       5://SYSTEM 5
           "CNV_ID_HMI" := "Settings_DB".ECnv_Sys[5].ID; // EXTRACTOR CONVEYOR
           "CNV_HMI".CNV2_Selected[5] := "CNV2_Selected";
           CASE "CNV_Level_Selected" OF
               1: //LEVEL 1
                   IF "CNV2_Selected" = 1 THEN
                       "CNV_ID_HMI(1)" := "Settings_DB".LCnv_Sys[5].Cnv_Level[1].Cnv1.ID; //CNV 1
                   ELSIF "CNV2_Selected" = 2 THEN
                       "CNV_ID_HMI(1)" := "Settings_DB".LCnv_Sys[5].Cnv_Level[1].Cnv2.ID; //CNV 2
                   END_IF;
               2: //LEVEL 2
                   IF "CNV2_Selected" = 1 THEN
                       "CNV_ID_HMI(1)" := "Settings_DB".LCnv_Sys[5].Cnv_Level[2].Cnv1.ID; //CNV 1
                   ELSIF "CNV2_Selected" = 2 THEN
                       "CNV_ID_HMI(1)" := "Settings_DB".LCnv_Sys[5].Cnv_Level[2].Cnv2.ID; //CNV 2
                   END_IF;
               3: //LEVEL 3
                   IF "CNV2_Selected" = 1 THEN
                       "CNV_ID_HMI(1)" := "Settings_DB".LCnv_Sys[5].Cnv_Level[3].Cnv1.ID; //CNV 1
                   ELSIF "CNV2_Selected" = 2 THEN
                       "CNV_ID_HMI(1)" := "Settings_DB".LCnv_Sys[5].Cnv_Level[3].Cnv2.ID; //CNV 2
                   END_IF;
               4: //LEVEL 4
                   IF "CNV2_Selected" = 1 THEN
                       "CNV_ID_HMI(1)" := "Settings_DB".LCnv_Sys[5].Cnv_Level[4].Cnv1.ID; //CNV 1
                   ELSIF "CNV2_Selected" = 2 THEN
                       "CNV_ID_HMI(1)" := "Settings_DB".LCnv_Sys[5].Cnv_Level[4].Cnv2.ID; //CNV 2
                   END_IF;
               5: //LEVEL 5
                   IF "CNV2_Selected" = 1 THEN
                       "CNV_ID_HMI(1)" := "Settings_DB".LCnv_Sys[5].Cnv_Level[5].Cnv1.ID; //CNV 1
                   ELSIF "CNV2_Selected" = 2 THEN
                       "CNV_ID_HMI(1)" := "Settings_DB".LCnv_Sys[5].Cnv_Level[5].Cnv2.ID; //CNV 2
                   END_IF;
               6: //LEVEL 6
                   IF "CNV2_Selected" = 1 THEN
                       "CNV_ID_HMI(1)" := "Settings_DB".LCnv_Sys[5].Cnv_Level[6].Cnv1.ID; //CNV 1
                   ELSIF "CNV2_Selected" = 2 THEN
                       "CNV_ID_HMI(1)" := "Settings_DB".LCnv_Sys[5].Cnv_Level[6].Cnv2.ID; //CNV 2
                   END_IF;
               7: //LEVEL 7
                   IF "CNV2_Selected" = 1 THEN
                       "CNV_ID_HMI(1)" := "Settings_DB".LCnv_Sys[5].Cnv_Level[7].Cnv1.ID; //CNV 1
                   ELSIF "CNV2_Selected" = 2 THEN
                       "CNV_ID_HMI(1)" := "Settings_DB".LCnv_Sys[5].Cnv_Level[7].Cnv2.ID; //CNV 2
                   END_IF;
               8: //LEVEL 8
                   IF "CNV2_Selected" = 1 THEN
                       "CNV_ID_HMI(1)" := "Settings_DB".LCnv_Sys[5].Cnv_Level[8].Cnv1.ID; //CNV 1
                   ELSIF "CNV2_Selected" = 2 THEN
                       "CNV_ID_HMI(1)" := "Settings_DB".LCnv_Sys[5].Cnv_Level[8].Cnv2.ID; //CNV 2
                   END_IF;
           END_CASE;
   END_CASE;
END_FUNCTION

FUNCTION "CNV_Selector_1" : Void   // FC60, SCL
{ S7_Optimized_Access := 'TRUE' }
VERSION : 0.1
// stored: AutoNumber true, IsIECCheckEnabled false, SetENOAutomatically false, UDAEnableTagReadback false
   VAR_INPUT
      Sys_No : UInt;
      Zone : UInt;
      CNV1_2_Selected : UInt;
   END_VAR
   VAR_OUTPUT
      ID : DInt;
      "ID(1)" : DInt;
   END_VAR
BEGIN
   //CNV SCREEN SELECTION
   CASE #Sys_No OF
       0:
           #ID := 0;
           #"ID(1)" := 0;

       1://SYSTEM 1
           #ID := "Settings_DB".ECnv_Sys[1].ID; // EXTRACTOR CONVEYOR
           CASE #Zone OF
               11: //LEVEL 1
                   IF #CNV1_2_Selected = 1 THEN
                       #"ID(1)" := "Settings_DB".LCnv_Sys[1].Cnv_Level[1].Cnv1.ID; //CNV 1
                   ELSIF #CNV1_2_Selected = 2 THEN
                       #"ID(1)" := "Settings_DB".LCnv_Sys[1].Cnv_Level[1].Cnv2.ID; //CNV 2
                   END_IF;
               12: //LEVEL 2
                   IF #CNV1_2_Selected = 1 THEN
                       #"ID(1)" := "Settings_DB".LCnv_Sys[1].Cnv_Level[2].Cnv1.ID; //CNV 1
                   ELSIF #CNV1_2_Selected = 2 THEN
                       #"ID(1)" := "Settings_DB".LCnv_Sys[1].Cnv_Level[2].Cnv2.ID; //CNV 2
                   END_IF;
               13: //LEVEL 3
                   IF #CNV1_2_Selected = 1 THEN
                       #"ID(1)" := "Settings_DB".LCnv_Sys[1].Cnv_Level[3].Cnv1.ID; //CNV 1
                   ELSIF #CNV1_2_Selected = 2 THEN
                       #"ID(1)" := "Settings_DB".LCnv_Sys[1].Cnv_Level[3].Cnv2.ID; //CNV 2
                   END_IF;
               14: //LEVEL 4
                   IF #CNV1_2_Selected = 1 THEN
                       #"ID(1)" := "Settings_DB".LCnv_Sys[1].Cnv_Level[4].Cnv1.ID; //CNV 1
                   ELSIF #CNV1_2_Selected = 2 THEN
                       #"ID(1)" := "Settings_DB".LCnv_Sys[1].Cnv_Level[4].Cnv2.ID; //CNV 2
                   END_IF;
               15: //LEVEL 5
                   IF #CNV1_2_Selected = 1 THEN
                       #"ID(1)" := "Settings_DB".LCnv_Sys[1].Cnv_Level[5].Cnv1.ID; //CNV 1
                   ELSIF #CNV1_2_Selected = 2 THEN
                       #"ID(1)" := "Settings_DB".LCnv_Sys[1].Cnv_Level[5].Cnv2.ID; //CNV 2
                   END_IF;
               16: //LEVEL 6
                   IF #CNV1_2_Selected = 1 THEN
                       #"ID(1)" := "Settings_DB".LCnv_Sys[1].Cnv_Level[6].Cnv1.ID; //CNV 1
                   ELSIF #CNV1_2_Selected = 2 THEN
                       #"ID(1)" := "Settings_DB".LCnv_Sys[1].Cnv_Level[6].Cnv2.ID; //CNV 2
                   END_IF;
               17: //LEVEL 7
                   IF #CNV1_2_Selected = 1 THEN
                       #"ID(1)" := "Settings_DB".LCnv_Sys[1].Cnv_Level[7].Cnv1.ID; //CNV 1
                   ELSIF #CNV1_2_Selected = 2 THEN
                       #"ID(1)" := "Settings_DB".LCnv_Sys[1].Cnv_Level[7].Cnv2.ID; //CNV 2
                   END_IF;
               18: //LEVEL 8
                   IF #CNV1_2_Selected = 1 THEN
                       #"ID(1)" := "Settings_DB".LCnv_Sys[1].Cnv_Level[8].Cnv1.ID; //CNV 1
                   ELSIF #CNV1_2_Selected = 2 THEN
                       #"ID(1)" := "Settings_DB".LCnv_Sys[1].Cnv_Level[8].Cnv2.ID; //CNV 2
                   END_IF;
               19: //LEVEL 1
                   IF #CNV1_2_Selected = 1 THEN
                       #"ID(1)" := "Settings_DB".LCnv_Sys[1].Cnv_Level[1].Cnv1.ID; //CNV 1
                   ELSIF #CNV1_2_Selected = 2 THEN
                       #"ID(1)" := "Settings_DB".LCnv_Sys[1].Cnv_Level[1].Cnv2.ID; //CNV 2
                   END_IF;
           END_CASE;

       2://SYSTEM 2
           #ID := "Settings_DB".ECnv_Sys[2].ID; // EXTRACTOR CONVEYOR
           CASE #Zone OF
               21: //LEVEL 1
                   IF #CNV1_2_Selected = 1 THEN
                       #"ID(1)" := "Settings_DB".LCnv_Sys[2].Cnv_Level[1].Cnv1.ID; //CNV 1
                   ELSIF #CNV1_2_Selected = 2 THEN
                       #"ID(1)" := "Settings_DB".LCnv_Sys[2].Cnv_Level[1].Cnv2.ID; //CNV 2
                   END_IF;
               22: //LEVEL 2
                   IF #CNV1_2_Selected = 1 THEN
                       #"ID(1)" := "Settings_DB".LCnv_Sys[2].Cnv_Level[2].Cnv1.ID; //CNV 1
                   ELSIF #CNV1_2_Selected = 2 THEN
                       #"ID(1)" := "Settings_DB".LCnv_Sys[2].Cnv_Level[2].Cnv2.ID; //CNV 2
                   END_IF;
               23: //LEVEL 3
                   IF #CNV1_2_Selected = 1 THEN
                       #"ID(1)" := "Settings_DB".LCnv_Sys[2].Cnv_Level[3].Cnv1.ID; //CNV 1
                   ELSIF #CNV1_2_Selected = 2 THEN
                       #"ID(1)" := "Settings_DB".LCnv_Sys[2].Cnv_Level[3].Cnv2.ID; //CNV 2
                   END_IF;
               24: //LEVEL 4
                   IF #CNV1_2_Selected = 1 THEN
                       #"ID(1)" := "Settings_DB".LCnv_Sys[2].Cnv_Level[4].Cnv1.ID; //CNV 1
                   ELSIF #CNV1_2_Selected = 2 THEN
                       #"ID(1)" := "Settings_DB".LCnv_Sys[2].Cnv_Level[4].Cnv2.ID; //CNV 2
                   END_IF;
               25: //LEVEL 5
                   IF #CNV1_2_Selected = 1 THEN
                       #"ID(1)" := "Settings_DB".LCnv_Sys[2].Cnv_Level[5].Cnv1.ID; //CNV 1
                   ELSIF #CNV1_2_Selected = 2 THEN
                       #"ID(1)" := "Settings_DB".LCnv_Sys[2].Cnv_Level[5].Cnv2.ID; //CNV 2
                   END_IF;
               26: //LEVEL 6
                   IF #CNV1_2_Selected = 1 THEN
                       #"ID(1)" := "Settings_DB".LCnv_Sys[2].Cnv_Level[6].Cnv1.ID; //CNV 1
                   ELSIF #CNV1_2_Selected = 2 THEN
                       #"ID(1)" := "Settings_DB".LCnv_Sys[2].Cnv_Level[6].Cnv2.ID; //CNV 2
                   END_IF;
               27: //LEVEL 7
                   IF #CNV1_2_Selected = 1 THEN
                       #"ID(1)" := "Settings_DB".LCnv_Sys[2].Cnv_Level[7].Cnv1.ID; //CNV 1
                   ELSIF #CNV1_2_Selected = 2 THEN
                       #"ID(1)" := "Settings_DB".LCnv_Sys[2].Cnv_Level[7].Cnv2.ID; //CNV 2
                   END_IF;
               28: //LEVEL 8
                   IF #CNV1_2_Selected = 1 THEN
                       #"ID(1)" := "Settings_DB".LCnv_Sys[2].Cnv_Level[8].Cnv1.ID; //CNV 1
                   ELSIF #CNV1_2_Selected = 2 THEN
                       #"ID(1)" := "Settings_DB".LCnv_Sys[2].Cnv_Level[8].Cnv2.ID; //CNV 2
                   END_IF;
               29: //LEVEL 1
                   IF #CNV1_2_Selected = 1 THEN
                       #"ID(1)" := "Settings_DB".LCnv_Sys[2].Cnv_Level[1].Cnv1.ID; //CNV 1
                   ELSIF #CNV1_2_Selected = 2 THEN
                       #"ID(1)" := "Settings_DB".LCnv_Sys[2].Cnv_Level[1].Cnv2.ID; //CNV 2
                   END_IF;
           END_CASE;

       3://SYSTEM 3
           #ID := "Settings_DB".ECnv_Sys[3].ID; // EXTRACTOR CONVEYOR
           CASE #Zone OF
               31: //LEVEL 1
                   IF #CNV1_2_Selected = 1 THEN
                       #"ID(1)" := "Settings_DB".LCnv_Sys[3].Cnv_Level[1].Cnv1.ID; //CNV 1
                   ELSIF #CNV1_2_Selected = 2 THEN
                       #"ID(1)" := "Settings_DB".LCnv_Sys[3].Cnv_Level[1].Cnv2.ID; //CNV 2
                   END_IF;
               32: //LEVEL 2
                   IF #CNV1_2_Selected = 1 THEN
                       #"ID(1)" := "Settings_DB".LCnv_Sys[3].Cnv_Level[2].Cnv1.ID; //CNV 1
                   ELSIF #CNV1_2_Selected = 2 THEN
                       #"ID(1)" := "Settings_DB".LCnv_Sys[3].Cnv_Level[2].Cnv2.ID; //CNV 2
                   END_IF;
               33: //LEVEL 3
                   IF #CNV1_2_Selected = 1 THEN
                       #"ID(1)" := "Settings_DB".LCnv_Sys[3].Cnv_Level[3].Cnv1.ID; //CNV 1
                   ELSIF #CNV1_2_Selected = 2 THEN
                       #"ID(1)" := "Settings_DB".LCnv_Sys[3].Cnv_Level[3].Cnv2.ID; //CNV 2
                   END_IF;
               34: //LEVEL 4
                   IF #CNV1_2_Selected = 1 THEN
                       #"ID(1)" := "Settings_DB".LCnv_Sys[3].Cnv_Level[4].Cnv1.ID; //CNV 1
                   ELSIF #CNV1_2_Selected = 2 THEN
                       #"ID(1)" := "Settings_DB".LCnv_Sys[3].Cnv_Level[4].Cnv2.ID; //CNV 2
                   END_IF;
               35: //LEVEL 5
                   IF #CNV1_2_Selected = 1 THEN
                       #"ID(1)" := "Settings_DB".LCnv_Sys[3].Cnv_Level[5].Cnv1.ID; //CNV 1
                   ELSIF #CNV1_2_Selected = 2 THEN
                       #"ID(1)" := "Settings_DB".LCnv_Sys[3].Cnv_Level[5].Cnv2.ID; //CNV 2
                   END_IF;
               36: //LEVEL 6
                   IF #CNV1_2_Selected = 1 THEN
                       #"ID(1)" := "Settings_DB".LCnv_Sys[3].Cnv_Level[6].Cnv1.ID; //CNV 1
                   ELSIF #CNV1_2_Selected = 2 THEN
                       #"ID(1)" := "Settings_DB".LCnv_Sys[3].Cnv_Level[6].Cnv2.ID; //CNV 2
                   END_IF;
               37: //LEVEL 7
                   IF #CNV1_2_Selected = 1 THEN
                       #"ID(1)" := "Settings_DB".LCnv_Sys[3].Cnv_Level[7].Cnv1.ID; //CNV 1
                   ELSIF #CNV1_2_Selected = 2 THEN
                       #"ID(1)" := "Settings_DB".LCnv_Sys[3].Cnv_Level[7].Cnv2.ID; //CNV 2
                   END_IF;
               38: //LEVEL 8
                   IF #CNV1_2_Selected = 1 THEN
                       #"ID(1)" := "Settings_DB".LCnv_Sys[3].Cnv_Level[8].Cnv1.ID; //CNV 1
                   ELSIF #CNV1_2_Selected = 2 THEN
                       #"ID(1)" := "Settings_DB".LCnv_Sys[3].Cnv_Level[8].Cnv2.ID; //CNV 2
                   END_IF;
               39: //LEVEL 1
                   IF #CNV1_2_Selected = 1 THEN
                       #"ID(1)" := "Settings_DB".LCnv_Sys[3].Cnv_Level[1].Cnv1.ID; //CNV 1
                   ELSIF #CNV1_2_Selected = 2 THEN
                       #"ID(1)" := "Settings_DB".LCnv_Sys[3].Cnv_Level[1].Cnv2.ID; //CNV 2
                   END_IF;
           END_CASE;

       4://SYSTEM 4
           #ID := "Settings_DB".ECnv_Sys[4].ID; // EXTRACTOR CONVEYOR
           CASE #Zone OF
               41: //LEVEL 1
                   IF #CNV1_2_Selected = 1 THEN
                       #"ID(1)" := "Settings_DB".LCnv_Sys[4].Cnv_Level[1].Cnv1.ID; //CNV 1
                   ELSIF #CNV1_2_Selected = 2 THEN
                       #"ID(1)" := "Settings_DB".LCnv_Sys[4].Cnv_Level[1].Cnv2.ID; //CNV 2
                   END_IF;
               42: //LEVEL 2
                   IF #CNV1_2_Selected = 1 THEN
                       #"ID(1)" := "Settings_DB".LCnv_Sys[4].Cnv_Level[2].Cnv1.ID; //CNV 1
                   ELSIF #CNV1_2_Selected = 2 THEN
                       #"ID(1)" := "Settings_DB".LCnv_Sys[4].Cnv_Level[2].Cnv2.ID; //CNV 2
                   END_IF;
               43: //LEVEL 3
                   IF #CNV1_2_Selected = 1 THEN
                       #"ID(1)" := "Settings_DB".LCnv_Sys[4].Cnv_Level[3].Cnv1.ID; //CNV 1
                   ELSIF #CNV1_2_Selected = 2 THEN
                       #"ID(1)" := "Settings_DB".LCnv_Sys[4].Cnv_Level[3].Cnv2.ID; //CNV 2
                   END_IF;
               44: //LEVEL 4
                   IF #CNV1_2_Selected = 1 THEN
                       #"ID(1)" := "Settings_DB".LCnv_Sys[4].Cnv_Level[4].Cnv1.ID; //CNV 1
                   ELSIF #CNV1_2_Selected = 2 THEN
                       #"ID(1)" := "Settings_DB".LCnv_Sys[4].Cnv_Level[4].Cnv2.ID; //CNV 2
                   END_IF;
               45: //LEVEL 5
                   IF #CNV1_2_Selected = 1 THEN
                       #"ID(1)" := "Settings_DB".LCnv_Sys[4].Cnv_Level[5].Cnv1.ID; //CNV 1
                   ELSIF #CNV1_2_Selected = 2 THEN
                       #"ID(1)" := "Settings_DB".LCnv_Sys[4].Cnv_Level[5].Cnv2.ID; //CNV 2
                   END_IF;
               46: //LEVEL 6
                   IF #CNV1_2_Selected = 1 THEN
                       #"ID(1)" := "Settings_DB".LCnv_Sys[4].Cnv_Level[6].Cnv1.ID; //CNV 1
                   ELSIF #CNV1_2_Selected = 2 THEN
                       #"ID(1)" := "Settings_DB".LCnv_Sys[4].Cnv_Level[6].Cnv2.ID; //CNV 2
                   END_IF;
               47: //LEVEL 7
                   IF #CNV1_2_Selected = 1 THEN
                       #"ID(1)" := "Settings_DB".LCnv_Sys[4].Cnv_Level[7].Cnv1.ID; //CNV 1
                   ELSIF #CNV1_2_Selected = 2 THEN
                       #"ID(1)" := "Settings_DB".LCnv_Sys[4].Cnv_Level[7].Cnv2.ID; //CNV 2
                   END_IF;
               48: //LEVEL 8
                   IF #CNV1_2_Selected = 1 THEN
                       #"ID(1)" := "Settings_DB".LCnv_Sys[4].Cnv_Level[8].Cnv1.ID; //CNV 1
                   ELSIF #CNV1_2_Selected = 2 THEN
                       #"ID(1)" := "Settings_DB".LCnv_Sys[4].Cnv_Level[8].Cnv2.ID; //CNV 2
                   END_IF;
               49: //LEVEL 1
                   IF #CNV1_2_Selected = 1 THEN
                       #"ID(1)" := "Settings_DB".LCnv_Sys[4].Cnv_Level[1].Cnv1.ID; //CNV 1
                   ELSIF #CNV1_2_Selected = 2 THEN
                       #"ID(1)" := "Settings_DB".LCnv_Sys[4].Cnv_Level[1].Cnv2.ID; //CNV 2
                   END_IF;
           END_CASE;

       5://SYSTEM 5
           #ID := "Settings_DB".ECnv_Sys[5].ID; // EXTRACTOR CONVEYOR
           CASE #Zone OF
               51: //LEVEL 1
                   IF #CNV1_2_Selected = 1 THEN
                       #"ID(1)" := "Settings_DB".LCnv_Sys[5].Cnv_Level[1].Cnv1.ID; //CNV 1
                   ELSIF #CNV1_2_Selected = 2 THEN
                       #"ID(1)" := "Settings_DB".LCnv_Sys[5].Cnv_Level[1].Cnv2.ID; //CNV 2
                   END_IF;
               52: //LEVEL 2
                   IF #CNV1_2_Selected = 1 THEN
                       #"ID(1)" := "Settings_DB".LCnv_Sys[5].Cnv_Level[2].Cnv1.ID; //CNV 1
                   ELSIF #CNV1_2_Selected = 2 THEN
                       #"ID(1)" := "Settings_DB".LCnv_Sys[5].Cnv_Level[2].Cnv2.ID; //CNV 2
                   END_IF;
               53: //LEVEL 3
                   IF #CNV1_2_Selected = 1 THEN
                       #"ID(1)" := "Settings_DB".LCnv_Sys[5].Cnv_Level[3].Cnv1.ID; //CNV 1
                   ELSIF #CNV1_2_Selected = 2 THEN
                       #"ID(1)" := "Settings_DB".LCnv_Sys[5].Cnv_Level[3].Cnv2.ID; //CNV 2
                   END_IF;
               54: //LEVEL 4
                   IF #CNV1_2_Selected = 1 THEN
                       #"ID(1)" := "Settings_DB".LCnv_Sys[5].Cnv_Level[4].Cnv1.ID; //CNV 1
                   ELSIF #CNV1_2_Selected = 2 THEN
                       #"ID(1)" := "Settings_DB".LCnv_Sys[5].Cnv_Level[4].Cnv2.ID; //CNV 2
                   END_IF;
               55: //LEVEL 5
                   IF #CNV1_2_Selected = 1 THEN
                       #"ID(1)" := "Settings_DB".LCnv_Sys[5].Cnv_Level[5].Cnv1.ID; //CNV 1
                   ELSIF #CNV1_2_Selected = 2 THEN
                       #"ID(1)" := "Settings_DB".LCnv_Sys[5].Cnv_Level[5].Cnv2.ID; //CNV 2
                   END_IF;
               56: //LEVEL 6
                   IF #CNV1_2_Selected = 1 THEN
                       #"ID(1)" := "Settings_DB".LCnv_Sys[5].Cnv_Level[6].Cnv1.ID; //CNV 1
                   ELSIF #CNV1_2_Selected = 2 THEN
                       #"ID(1)" := "Settings_DB".LCnv_Sys[5].Cnv_Level[6].Cnv2.ID; //CNV 2
                   END_IF;
               57: //LEVEL 7
                   IF #CNV1_2_Selected = 1 THEN
                       #"ID(1)" := "Settings_DB".LCnv_Sys[5].Cnv_Level[7].Cnv1.ID; //CNV 1
                   ELSIF #CNV1_2_Selected = 2 THEN
                       #"ID(1)" := "Settings_DB".LCnv_Sys[5].Cnv_Level[7].Cnv2.ID; //CNV 2
                   END_IF;
               58: //LEVEL 8
                   IF #CNV1_2_Selected = 1 THEN
                       #"ID(1)" := "Settings_DB".LCnv_Sys[5].Cnv_Level[8].Cnv1.ID; //CNV 1
                   ELSIF #CNV1_2_Selected = 2 THEN
                       #"ID(1)" := "Settings_DB".LCnv_Sys[5].Cnv_Level[8].Cnv2.ID; //CNV 2
                   END_IF;
               59: //LEVEL 1
                   IF #CNV1_2_Selected = 1 THEN
                       #"ID(1)" := "Settings_DB".LCnv_Sys[5].Cnv_Level[1].Cnv1.ID; //CNV 1
                   ELSIF #CNV1_2_Selected = 2 THEN
                       #"ID(1)" := "Settings_DB".LCnv_Sys[5].Cnv_Level[1].Cnv2.ID; //CNV 2
                   END_IF;
           END_CASE;
   END_CASE;
END_FUNCTION

FUNCTION "CharsArrayToString" : String   // FC27, SCL
{ S7_Optimized_Access := 'TRUE' }
VERSION : 0.1
// stored: AutoNumber true, IsIECCheckEnabled false, SetENOAutomatically false, UDAEnableTagReadback false
   VAR_INPUT
      Lenght : Int;
      CharsArray : Array[1..16] of Char;
   END_VAR
   VAR_TEMP
      tempStr_1 : String;
      foundPos : Int;
      i : Int;
   END_VAR
BEGIN
   #tempStr_1 := '';
   FOR #i := 1 TO MIN(IN1 := #Lenght - 1, IN2 := 16) DO
       IF #CharsArray[#i] <> '$00' THEN
           #tempStr_1 := CONCAT(IN1 := #tempStr_1, IN2 := CHAR_TO_STRING(#CharsArray[#i]));
       END_IF;
   END_FOR;

   // Remove '$00'
   // string 1
   #foundPos := FIND(IN1 := #tempStr_1, IN2 := '$00');
   WHILE #foundPos > 0 DO
       #tempStr_1 := REPLACE(IN1 := #tempStr_1, IN2 := '', P := #foundPos, L := 1);
       #foundPos := FIND(IN1 := #tempStr_1, IN2 := '$00');
   END_WHILE;

   #CharsArrayToString := #tempStr_1;
END_FUNCTION

FUNCTION_BLOCK "Conveyor_HMI_FB"   // FB20, SCL
{ S7_Optimized_Access := 'TRUE' }
VERSION : 0.1
// stored: AutoNumber true, IsIECCheckEnabled false, IsRetainMemResEnabled false, MemoryReserve 100, SetENOAutomatically false, UDAEnableTagReadback false
   VAR
      R_Charge_Cnv_Commands { S7_SetPoint := 'True'} : R_TRIG;
      T_Reset_Charge { S7_SetPoint := 'True'} : TON_TIME;
   END_VAR
   VAR_TEMP
      i : UInt;
      J : UInt;
      No_Light_Guard : Bool;
   END_VAR
BEGIN
   "CNV_Selector"();

   REGION SEND/RECEIVE BUTTON
       IF "CNV_System_Selected" = 1 AND NOT "Control_DB".VTD_Sys[1].Running AND "Control_DB".VTD_Sys[1].Current_Level <> 0 THEN
           IF "CNV2_Selected" = 1 AND "HMI_DB".ScreenNo_Main = 2 THEN
               //CNV 1
               IF "Control_DB".ECnv_Sys[1].Cnv_Occupied AND NOT "Control_DB".LCnv_Sys[1].Cnv_Level["Control_DB".VTD_Sys[1].Current_Level].Cnv1.Cnv_Occupied AND
                   NOT "Control_DB".ECnv_Sys[1].Running AND NOT "Control_DB".LCnv_Sys[1].Cnv_Level["Control_DB".VTD_Sys[1].Current_Level].Cnv1.Running AND
                   "Control_DB".LCnv_Sys[1].Cnv_Level["Control_DB".VTD_Sys[1].Current_Level].Cnv1.Pallet_Type <> 1 AND "Control_DB".ECnv_Sys[1].Pallet_Type <> 5 THEN
                   "CNV_HMI".In_Out[1] := TRUE;
                   "CNV_In_Out" := TRUE;
               ELSIF NOT "Control_DB".ECnv_Sys[1].Cnv_Occupied AND "Control_DB".LCnv_Sys[1].Cnv_Level["Control_DB".VTD_Sys[1].Current_Level].Cnv1.Cnv_Occupied AND
                   NOT "Control_DB".ECnv_Sys[1].Running AND NOT "Control_DB".LCnv_Sys[1].Cnv_Level["Control_DB".VTD_Sys[1].Current_Level].Cnv1.Running THEN
                   "CNV_HMI".In_Out[1] := FALSE;
                   "CNV_In_Out" := FALSE;
               ELSE
                   ;
               END_IF;
               //CNV 2
           ELSIF "CNV2_Selected" = 2 AND "HMI_DB".ScreenNo_Main = 2 THEN   //CNV 2
               IF "Control_DB".ECnv_Sys[1].Cnv_Occupied AND NOT "Control_DB".LCnv_Sys[1].Cnv_Level["Control_DB".VTD_Sys[1].Current_Level].Cnv2.Cnv_Occupied AND
                   NOT "Control_DB".ECnv_Sys[1].Running AND NOT "Control_DB".LCnv_Sys[1].Cnv_Level["Control_DB".VTD_Sys[1].Current_Level].Cnv2.Running AND
                   "Control_DB".LCnv_Sys[1].Cnv_Level["Control_DB".VTD_Sys[1].Current_Level].Cnv2.Pallet_Type <> 1 AND "Control_DB".ECnv_Sys[1].Pallet_Type <> 5 THEN
                   "CNV_HMI".In_Out[1] := TRUE;
                   "CNV_In_Out" := TRUE;
               ELSIF NOT "Control_DB".ECnv_Sys[1].Cnv_Occupied AND "Control_DB".LCnv_Sys[1].Cnv_Level["Control_DB".VTD_Sys[1].Current_Level].Cnv2.Cnv_Occupied AND
                   NOT "Control_DB".ECnv_Sys[1].Running AND NOT "Control_DB".LCnv_Sys[1].Cnv_Level["Control_DB".VTD_Sys[1].Current_Level].Cnv2.Running THEN
                   "CNV_HMI".In_Out[1] := FALSE;
                   "CNV_In_Out" := FALSE;
               ELSE
                   ;
               END_IF;
           END_IF;
       END_IF;

       IF "CNV_System_Selected" = 2 AND NOT "Control_DB".VTD_Sys[2].Running AND "Control_DB".VTD_Sys[2].Current_Level <> 0 THEN
           IF "CNV2_Selected" = 1 AND "HMI_DB".ScreenNo_Main = 2 THEN
               //CNV 1
               IF "Control_DB".ECnv_Sys[2].Cnv_Occupied AND NOT "Control_DB".LCnv_Sys[2].Cnv_Level["Control_DB".VTD_Sys[2].Current_Level].Cnv1.Cnv_Occupied AND
                   NOT "Control_DB".ECnv_Sys[2].Running AND NOT "Control_DB".LCnv_Sys[2].Cnv_Level["Control_DB".VTD_Sys[2].Current_Level].Cnv1.Running AND
                   "Control_DB".LCnv_Sys[2].Cnv_Level["Control_DB".VTD_Sys[2].Current_Level].Cnv1.Pallet_Type <> 1 AND "Control_DB".ECnv_Sys[2].Pallet_Type <> 5 THEN
                   "CNV_HMI".In_Out[2] := TRUE;
                   "CNV_In_Out" := TRUE;
               ELSIF NOT "Control_DB".ECnv_Sys[2].Cnv_Occupied AND "Control_DB".LCnv_Sys[2].Cnv_Level["Control_DB".VTD_Sys[2].Current_Level].Cnv1.Cnv_Occupied AND
                   NOT "Control_DB".ECnv_Sys[2].Running AND NOT "Control_DB".LCnv_Sys[2].Cnv_Level["Control_DB".VTD_Sys[2].Current_Level].Cnv1.Running THEN
                   "CNV_HMI".In_Out[2] := FALSE;
                   "CNV_In_Out" := FALSE;
               ELSE
                   ;
               END_IF;
               //CNV 2
           ELSIF "CNV2_Selected" = 2 AND "HMI_DB".ScreenNo_Main = 2 THEN   //CNV 2
               IF "Control_DB".ECnv_Sys[2].Cnv_Occupied AND NOT "Control_DB".LCnv_Sys[2].Cnv_Level["Control_DB".VTD_Sys[2].Current_Level].Cnv2.Cnv_Occupied AND
                   NOT "Control_DB".ECnv_Sys[2].Running AND NOT "Control_DB".LCnv_Sys[2].Cnv_Level["Control_DB".VTD_Sys[2].Current_Level].Cnv2.Running AND
                   "Control_DB".LCnv_Sys[2].Cnv_Level["Control_DB".VTD_Sys[2].Current_Level].Cnv2.Pallet_Type <> 1 AND "Control_DB".ECnv_Sys[2].Pallet_Type <> 5 THEN
                   "CNV_HMI".In_Out[2] := TRUE;
                   "CNV_In_Out" := TRUE;
               ELSIF NOT "Control_DB".ECnv_Sys[2].Cnv_Occupied AND "Control_DB".LCnv_Sys[2].Cnv_Level["Control_DB".VTD_Sys[2].Current_Level].Cnv2.Cnv_Occupied AND
                   NOT "Control_DB".ECnv_Sys[2].Running AND NOT "Control_DB".LCnv_Sys[2].Cnv_Level["Control_DB".VTD_Sys[2].Current_Level].Cnv2.Running THEN
                   "CNV_HMI".In_Out[2] := FALSE;
                   "CNV_In_Out" := FALSE;
               ELSE
                   ;
               END_IF;
           END_IF;
       END_IF;

       IF "CNV_System_Selected" = 3 AND NOT "Control_DB".VTD_Sys[3].Running AND "Control_DB".VTD_Sys[3].Current_Level <> 0 THEN
           IF "CNV2_Selected" = 1 AND "HMI_DB".ScreenNo_Main = 2 THEN
               //CNV 1
               IF "Control_DB".ECnv_Sys[3].Cnv_Occupied AND NOT "Control_DB".LCnv_Sys[3].Cnv_Level["Control_DB".VTD_Sys[3].Current_Level].Cnv1.Cnv_Occupied AND
                   NOT "Control_DB".ECnv_Sys[3].Running AND NOT "Control_DB".LCnv_Sys[3].Cnv_Level["Control_DB".VTD_Sys[3].Current_Level].Cnv1.Running THEN
                   "CNV_HMI".In_Out[3] := TRUE;
                   "CNV_In_Out" := TRUE;
               ELSIF NOT "Control_DB".ECnv_Sys[3].Cnv_Occupied AND "Control_DB".LCnv_Sys[3].Cnv_Level["Control_DB".VTD_Sys[3].Current_Level].Cnv1.Cnv_Occupied AND
                   NOT "Control_DB".ECnv_Sys[3].Running AND NOT "Control_DB".LCnv_Sys[3].Cnv_Level["Control_DB".VTD_Sys[3].Current_Level].Cnv1.Running THEN
                   "CNV_HMI".In_Out[3] := FALSE;
                   "CNV_In_Out" := FALSE;
               ELSE
                   ;
               END_IF;
               //CNV 2
           ELSIF "CNV2_Selected" = 2 AND "HMI_DB".ScreenNo_Main = 2 THEN   //CNV 2
               IF "Control_DB".ECnv_Sys[3].Cnv_Occupied AND NOT "Control_DB".LCnv_Sys[3].Cnv_Level["Control_DB".VTD_Sys[3].Current_Level].Cnv2.Cnv_Occupied AND
                   NOT "Control_DB".ECnv_Sys[3].Running AND NOT "Control_DB".LCnv_Sys[3].Cnv_Level["Control_DB".VTD_Sys[3].Current_Level].Cnv2.Running THEN
                   "CNV_HMI".In_Out[3] := TRUE;
                   "CNV_In_Out" := TRUE;
               ELSIF NOT "Control_DB".ECnv_Sys[3].Cnv_Occupied AND "Control_DB".LCnv_Sys[3].Cnv_Level["Control_DB".VTD_Sys[3].Current_Level].Cnv2.Cnv_Occupied AND
                   NOT "Control_DB".ECnv_Sys[3].Running AND NOT "Control_DB".LCnv_Sys[3].Cnv_Level["Control_DB".VTD_Sys[3].Current_Level].Cnv2.Running THEN
                   "CNV_HMI".In_Out[3] := FALSE;
                   "CNV_In_Out" := FALSE;
               ELSE
                   ;
               END_IF;
           END_IF;
       END_IF;

       IF "CNV_System_Selected" = 4 AND NOT "Control_DB".VTD_Sys[4].Running AND "Control_DB".VTD_Sys[4].Current_Level <> 0 THEN
           IF "CNV2_Selected" = 1 AND "HMI_DB".ScreenNo_Main = 2 THEN
               //CNV 1
               IF "Control_DB".ECnv_Sys[4].Cnv_Occupied AND NOT "Control_DB".LCnv_Sys[4].Cnv_Level["Control_DB".VTD_Sys[4].Current_Level].Cnv1.Cnv_Occupied AND
                   NOT "Control_DB".ECnv_Sys[4].Running AND NOT "Control_DB".LCnv_Sys[4].Cnv_Level["Control_DB".VTD_Sys[4].Current_Level].Cnv1.Running THEN
                   "CNV_HMI".In_Out[4] := TRUE;
                   "CNV_In_Out" := TRUE;
               ELSIF NOT "Control_DB".ECnv_Sys[4].Cnv_Occupied AND "Control_DB".LCnv_Sys[4].Cnv_Level["Control_DB".VTD_Sys[4].Current_Level].Cnv1.Cnv_Occupied AND
                   NOT "Control_DB".ECnv_Sys[4].Running AND NOT "Control_DB".LCnv_Sys[4].Cnv_Level["Control_DB".VTD_Sys[4].Current_Level].Cnv1.Running THEN
                   "CNV_HMI".In_Out[4] := FALSE;
                   "CNV_In_Out" := FALSE;
               ELSE
                   ;
               END_IF;
           END_IF;
       END_IF;

       IF "CNV_System_Selected" = 5 AND NOT "Control_DB".VTD_Sys[5].Running AND "Control_DB".VTD_Sys[5].Current_Level <> 0 THEN
           IF "CNV2_Selected" = 1 AND "HMI_DB".ScreenNo_Main = 2 THEN
               //CNV 1
               IF "Control_DB".ECnv_Sys[5].Cnv_Occupied AND NOT "Control_DB".LCnv_Sys[5].Cnv_Level["Control_DB".VTD_Sys[5].Current_Level].Cnv1.Cnv_Occupied AND
                   NOT "Control_DB".ECnv_Sys[5].Running AND NOT "Control_DB".LCnv_Sys[5].Cnv_Level["Control_DB".VTD_Sys[5].Current_Level].Cnv1.Running THEN
                   "CNV_HMI".In_Out[5] := TRUE;
                   "CNV_In_Out" := TRUE;
               ELSIF NOT "Control_DB".ECnv_Sys[5].Cnv_Occupied AND "Control_DB".LCnv_Sys[5].Cnv_Level["Control_DB".VTD_Sys[5].Current_Level].Cnv1.Cnv_Occupied AND
                   NOT "Control_DB".ECnv_Sys[5].Running AND NOT "Control_DB".LCnv_Sys[5].Cnv_Level["Control_DB".VTD_Sys[5].Current_Level].Cnv1.Running THEN
                   "CNV_HMI".In_Out[5] := FALSE;
                   "CNV_In_Out" := FALSE;
               ELSE
                   ;
               END_IF;
           END_IF;
       END_IF;
   END_REGION ;

   REGION Assign Conveyor 1
       REGION CHARGE DATA FROM THE CORRECT CONVEYOR
           //CHARGE DATA CHANGING CONVEYORS ID
           IF "CNV_ID_HMI" <> "CNV_ID_HMI_Old" THEN
               "Screen_DB".Charge_Cnv_Commands := TRUE;
               "CNV_ID_HMI_Old" := "CNV_ID_HMI";
           END_IF;
           #R_Charge_Cnv_Commands(CLK := "Screen_DB".Charge_Cnv_Commands OR "HMI_DB".ScreenNo_Main = 2);

           //CHARGE ONCE THE COMMANDS STATUS
           IF "Screen_DB".Charge_Cnv_Commands THEN
               CASE "CNV_ID_HMI" OF
                       //SYSTEM 1
                   120001:
                       "Enable_HMI" := "Control_DB".ECnv_Sys[1].Instruction.Enable;
                       "Mode_Change_HMI" := "Control_DB".ECnv_Sys[1].Instruction.Mode_Change;
                       "Task_ID_HMI" := "Control_DB".ECnv_Sys[1].Instruction.Task_ID;
                       "Transfer_To_ID_HMI" := "Control_DB".ECnv_Sys[1].Instruction.Transfer_To_ID;
                       "Transfer_From_ID_HMI" := "Control_DB".ECnv_Sys[1].Instruction.Transfer_From_ID;
                       "Pallet_Allignment_HMI" := "Control_DB".ECnv_Sys[1].Instruction.Pallet_Allignment;
                   120101:
                       "Enable_HMI" := "Control_DB".ECnv_Sys[1].Instruction.Enable;
                       "Mode_Change_HMI" := "Control_DB".ECnv_Sys[1].Instruction.Mode_Change;
                       "Task_ID_HMI" := "Control_DB".ECnv_Sys[1].Instruction.Task_ID;
                       "Transfer_To_ID_HMI" := "Control_DB".ECnv_Sys[1].Instruction.Transfer_To_ID;
                       "Transfer_From_ID_HMI" := "Control_DB".ECnv_Sys[1].Instruction.Transfer_From_ID;
                       "Pallet_Allignment_HMI" := "Control_DB".ECnv_Sys[1].Instruction.Pallet_Allignment;
                   120201:
                       "Enable_HMI" := "Control_DB".ECnv_Sys[1].Instruction.Enable;
                       "Mode_Change_HMI" := "Control_DB".ECnv_Sys[1].Instruction.Mode_Change;
                       "Task_ID_HMI" := "Control_DB".ECnv_Sys[1].Instruction.Task_ID;
                       "Transfer_To_ID_HMI" := "Control_DB".ECnv_Sys[1].Instruction.Transfer_To_ID;
                       "Transfer_From_ID_HMI" := "Control_DB".ECnv_Sys[1].Instruction.Transfer_From_ID;
                       "Pallet_Allignment_HMI" := "Control_DB".ECnv_Sys[1].Instruction.Pallet_Allignment;
                   120301:
                       "Enable_HMI" := "Control_DB".ECnv_Sys[1].Instruction.Enable;
                       "Mode_Change_HMI" := "Control_DB".ECnv_Sys[1].Instruction.Mode_Change;
                       "Task_ID_HMI" := "Control_DB".ECnv_Sys[1].Instruction.Task_ID;
                       "Transfer_To_ID_HMI" := "Control_DB".ECnv_Sys[1].Instruction.Transfer_To_ID;
                       "Transfer_From_ID_HMI" := "Control_DB".ECnv_Sys[1].Instruction.Transfer_From_ID;
                       "Pallet_Allignment_HMI" := "Control_DB".ECnv_Sys[1].Instruction.Pallet_Allignment;
                   120401:
                       "Enable_HMI" := "Control_DB".ECnv_Sys[1].Instruction.Enable;
                       "Mode_Change_HMI" := "Control_DB".ECnv_Sys[1].Instruction.Mode_Change;
                       "Task_ID_HMI" := "Control_DB".ECnv_Sys[1].Instruction.Task_ID;
                       "Transfer_To_ID_HMI" := "Control_DB".ECnv_Sys[1].Instruction.Transfer_To_ID;
                       "Transfer_From_ID_HMI" := "Control_DB".ECnv_Sys[1].Instruction.Transfer_From_ID;
                       "Pallet_Allignment_HMI" := "Control_DB".ECnv_Sys[1].Instruction.Pallet_Allignment;
                   120501:
                       "Enable_HMI" := "Control_DB".ECnv_Sys[1].Instruction.Enable;
                       "Mode_Change_HMI" := "Control_DB".ECnv_Sys[1].Instruction.Mode_Change;
                       "Task_ID_HMI" := "Control_DB".ECnv_Sys[1].Instruction.Task_ID;
                       "Transfer_To_ID_HMI" := "Control_DB".ECnv_Sys[1].Instruction.Transfer_To_ID;
                       "Transfer_From_ID_HMI" := "Control_DB".ECnv_Sys[1].Instruction.Transfer_From_ID;
                       "Pallet_Allignment_HMI" := "Control_DB".ECnv_Sys[1].Instruction.Pallet_Allignment;
                   120601:
                       "Enable_HMI" := "Control_DB".ECnv_Sys[1].Instruction.Enable;
                       "Mode_Change_HMI" := "Control_DB".ECnv_Sys[1].Instruction.Mode_Change;
                       "Task_ID_HMI" := "Control_DB".ECnv_Sys[1].Instruction.Task_ID;
                       "Transfer_To_ID_HMI" := "Control_DB".ECnv_Sys[1].Instruction.Transfer_To_ID;
                       "Transfer_From_ID_HMI" := "Control_DB".ECnv_Sys[1].Instruction.Transfer_From_ID;
                       "Pallet_Allignment_HMI" := "Control_DB".ECnv_Sys[1].Instruction.Pallet_Allignment;
                   120701:
                       "Enable_HMI" := "Control_DB".ECnv_Sys[1].Instruction.Enable;
                       "Mode_Change_HMI" := "Control_DB".ECnv_Sys[1].Instruction.Mode_Change;
                       "Task_ID_HMI" := "Control_DB".ECnv_Sys[1].Instruction.Task_ID;
                       "Transfer_To_ID_HMI" := "Control_DB".ECnv_Sys[1].Instruction.Transfer_To_ID;
                       "Transfer_From_ID_HMI" := "Control_DB".ECnv_Sys[1].Instruction.Transfer_From_ID;
                       "Pallet_Allignment_HMI" := "Control_DB".ECnv_Sys[1].Instruction.Pallet_Allignment;
                   120801:
                       "Enable_HMI" := "Control_DB".ECnv_Sys[1].Instruction.Enable;
                       "Mode_Change_HMI" := "Control_DB".ECnv_Sys[1].Instruction.Mode_Change;
                       "Task_ID_HMI" := "Control_DB".ECnv_Sys[1].Instruction.Task_ID;
                       "Transfer_To_ID_HMI" := "Control_DB".ECnv_Sys[1].Instruction.Transfer_To_ID;
                       "Transfer_From_ID_HMI" := "Control_DB".ECnv_Sys[1].Instruction.Transfer_From_ID;
                       "Pallet_Allignment_HMI" := "Control_DB".ECnv_Sys[1].Instruction.Pallet_Allignment;

                       //SYSTEM 2
                   120002:
                       "Enable_HMI" := "Control_DB".ECnv_Sys[2].Instruction.Enable;
                       "Mode_Change_HMI" := "Control_DB".ECnv_Sys[2].Instruction.Mode_Change;
                       "Task_ID_HMI" := "Control_DB".ECnv_Sys[2].Instruction.Task_ID;
                       "Transfer_To_ID_HMI" := "Control_DB".ECnv_Sys[2].Instruction.Transfer_To_ID;
                       "Transfer_From_ID_HMI" := "Control_DB".ECnv_Sys[2].Instruction.Transfer_From_ID;
                       "Pallet_Allignment_HMI" := "Control_DB".ECnv_Sys[2].Instruction.Pallet_Allignment;
                   120102:
                       "Enable_HMI" := "Control_DB".ECnv_Sys[2].Instruction.Enable;
                       "Mode_Change_HMI" := "Control_DB".ECnv_Sys[2].Instruction.Mode_Change;
                       "Task_ID_HMI" := "Control_DB".ECnv_Sys[2].Instruction.Task_ID;
                       "Transfer_To_ID_HMI" := "Control_DB".ECnv_Sys[2].Instruction.Transfer_To_ID;
                       "Transfer_From_ID_HMI" := "Control_DB".ECnv_Sys[2].Instruction.Transfer_From_ID;
                       "Pallet_Allignment_HMI" := "Control_DB".ECnv_Sys[2].Instruction.Pallet_Allignment;
                   120202:
                       "Enable_HMI" := "Control_DB".ECnv_Sys[2].Instruction.Enable;
                       "Mode_Change_HMI" := "Control_DB".ECnv_Sys[2].Instruction.Mode_Change;
                       "Task_ID_HMI" := "Control_DB".ECnv_Sys[2].Instruction.Task_ID;
                       "Transfer_To_ID_HMI" := "Control_DB".ECnv_Sys[2].Instruction.Transfer_To_ID;
                       "Transfer_From_ID_HMI" := "Control_DB".ECnv_Sys[2].Instruction.Transfer_From_ID;
                       "Pallet_Allignment_HMI" := "Control_DB".ECnv_Sys[2].Instruction.Pallet_Allignment;
                   120302:
                       "Enable_HMI" := "Control_DB".ECnv_Sys[2].Instruction.Enable;
                       "Mode_Change_HMI" := "Control_DB".ECnv_Sys[2].Instruction.Mode_Change;
                       "Task_ID_HMI" := "Control_DB".ECnv_Sys[2].Instruction.Task_ID;
                       "Transfer_To_ID_HMI" := "Control_DB".ECnv_Sys[2].Instruction.Transfer_To_ID;
                       "Transfer_From_ID_HMI" := "Control_DB".ECnv_Sys[2].Instruction.Transfer_From_ID;
                       "Pallet_Allignment_HMI" := "Control_DB".ECnv_Sys[2].Instruction.Pallet_Allignment;
                   120402:
                       "Enable_HMI" := "Control_DB".ECnv_Sys[2].Instruction.Enable;
                       "Mode_Change_HMI" := "Control_DB".ECnv_Sys[2].Instruction.Mode_Change;
                       "Task_ID_HMI" := "Control_DB".ECnv_Sys[2].Instruction.Task_ID;
                       "Transfer_To_ID_HMI" := "Control_DB".ECnv_Sys[2].Instruction.Transfer_To_ID;
                       "Transfer_From_ID_HMI" := "Control_DB".ECnv_Sys[2].Instruction.Transfer_From_ID;
                       "Pallet_Allignment_HMI" := "Control_DB".ECnv_Sys[2].Instruction.Pallet_Allignment;
                   120502:
                       "Enable_HMI" := "Control_DB".ECnv_Sys[2].Instruction.Enable;
                       "Mode_Change_HMI" := "Control_DB".ECnv_Sys[2].Instruction.Mode_Change;
                       "Task_ID_HMI" := "Control_DB".ECnv_Sys[2].Instruction.Task_ID;
                       "Transfer_To_ID_HMI" := "Control_DB".ECnv_Sys[2].Instruction.Transfer_To_ID;
                       "Transfer_From_ID_HMI" := "Control_DB".ECnv_Sys[2].Instruction.Transfer_From_ID;
                       "Pallet_Allignment_HMI" := "Control_DB".ECnv_Sys[2].Instruction.Pallet_Allignment;
                   120602:
                       "Enable_HMI" := "Control_DB".ECnv_Sys[2].Instruction.Enable;
                       "Mode_Change_HMI" := "Control_DB".ECnv_Sys[2].Instruction.Mode_Change;
                       "Task_ID_HMI" := "Control_DB".ECnv_Sys[2].Instruction.Task_ID;
                       "Transfer_To_ID_HMI" := "Control_DB".ECnv_Sys[2].Instruction.Transfer_To_ID;
                       "Transfer_From_ID_HMI" := "Control_DB".ECnv_Sys[2].Instruction.Transfer_From_ID;
                       "Pallet_Allignment_HMI" := "Control_DB".ECnv_Sys[2].Instruction.Pallet_Allignment;
                   120702:
                       "Enable_HMI" := "Control_DB".ECnv_Sys[2].Instruction.Enable;
                       "Mode_Change_HMI" := "Control_DB".ECnv_Sys[2].Instruction.Mode_Change;
                       "Task_ID_HMI" := "Control_DB".ECnv_Sys[2].Instruction.Task_ID;
                       "Transfer_To_ID_HMI" := "Control_DB".ECnv_Sys[2].Instruction.Transfer_To_ID;
                       "Transfer_From_ID_HMI" := "Control_DB".ECnv_Sys[2].Instruction.Transfer_From_ID;
                       "Pallet_Allignment_HMI" := "Control_DB".ECnv_Sys[2].Instruction.Pallet_Allignment;
                   120802:
                       "Enable_HMI" := "Control_DB".ECnv_Sys[2].Instruction.Enable;
                       "Mode_Change_HMI" := "Control_DB".ECnv_Sys[2].Instruction.Mode_Change;
                       "Task_ID_HMI" := "Control_DB".ECnv_Sys[2].Instruction.Task_ID;
                       "Transfer_To_ID_HMI" := "Control_DB".ECnv_Sys[2].Instruction.Transfer_To_ID;
                       "Transfer_From_ID_HMI" := "Control_DB".ECnv_Sys[2].Instruction.Transfer_From_ID;
                       "Pallet_Allignment_HMI" := "Control_DB".ECnv_Sys[2].Instruction.Pallet_Allignment;

                       //SYSTEM 3
                   120003:
                       "Enable_HMI" := "Control_DB".ECnv_Sys[3].Instruction.Enable;
                       "Mode_Change_HMI" := "Control_DB".ECnv_Sys[3].Instruction.Mode_Change;
                       "Task_ID_HMI" := "Control_DB".ECnv_Sys[3].Instruction.Task_ID;
                       "Transfer_To_ID_HMI" := "Control_DB".ECnv_Sys[3].Instruction.Transfer_To_ID;
                       "Transfer_From_ID_HMI" := "Control_DB".ECnv_Sys[3].Instruction.Transfer_From_ID;
                       "Pallet_Allignment_HMI" := "Control_DB".ECnv_Sys[3].Instruction.Pallet_Allignment;
                   120103:
                       "Enable_HMI" := "Control_DB".ECnv_Sys[3].Instruction.Enable;
                       "Mode_Change_HMI" := "Control_DB".ECnv_Sys[3].Instruction.Mode_Change;
                       "Task_ID_HMI" := "Control_DB".ECnv_Sys[3].Instruction.Task_ID;
                       "Transfer_To_ID_HMI" := "Control_DB".ECnv_Sys[3].Instruction.Transfer_To_ID;
                       "Transfer_From_ID_HMI" := "Control_DB".ECnv_Sys[3].Instruction.Transfer_From_ID;
                       "Pallet_Allignment_HMI" := "Control_DB".ECnv_Sys[3].Instruction.Pallet_Allignment;
                   120203:
                       "Enable_HMI" := "Control_DB".ECnv_Sys[3].Instruction.Enable;
                       "Mode_Change_HMI" := "Control_DB".ECnv_Sys[3].Instruction.Mode_Change;
                       "Task_ID_HMI" := "Control_DB".ECnv_Sys[3].Instruction.Task_ID;
                       "Transfer_To_ID_HMI" := "Control_DB".ECnv_Sys[3].Instruction.Transfer_To_ID;
                       "Transfer_From_ID_HMI" := "Control_DB".ECnv_Sys[3].Instruction.Transfer_From_ID;
                       "Pallet_Allignment_HMI" := "Control_DB".ECnv_Sys[3].Instruction.Pallet_Allignment;
                   120303:
                       "Enable_HMI" := "Control_DB".ECnv_Sys[3].Instruction.Enable;
                       "Mode_Change_HMI" := "Control_DB".ECnv_Sys[3].Instruction.Mode_Change;
                       "Task_ID_HMI" := "Control_DB".ECnv_Sys[3].Instruction.Task_ID;
                       "Transfer_To_ID_HMI" := "Control_DB".ECnv_Sys[3].Instruction.Transfer_To_ID;
                       "Transfer_From_ID_HMI" := "Control_DB".ECnv_Sys[3].Instruction.Transfer_From_ID;
                       "Pallet_Allignment_HMI" := "Control_DB".ECnv_Sys[3].Instruction.Pallet_Allignment;
                   120403:
                       "Enable_HMI" := "Control_DB".ECnv_Sys[3].Instruction.Enable;
                       "Mode_Change_HMI" := "Control_DB".ECnv_Sys[3].Instruction.Mode_Change;
                       "Task_ID_HMI" := "Control_DB".ECnv_Sys[3].Instruction.Task_ID;
                       "Transfer_To_ID_HMI" := "Control_DB".ECnv_Sys[3].Instruction.Transfer_To_ID;
                       "Transfer_From_ID_HMI" := "Control_DB".ECnv_Sys[3].Instruction.Transfer_From_ID;
                       "Pallet_Allignment_HMI" := "Control_DB".ECnv_Sys[3].Instruction.Pallet_Allignment;
                   120503:
                       "Enable_HMI" := "Control_DB".ECnv_Sys[3].Instruction.Enable;
                       "Mode_Change_HMI" := "Control_DB".ECnv_Sys[3].Instruction.Mode_Change;
                       "Task_ID_HMI" := "Control_DB".ECnv_Sys[3].Instruction.Task_ID;
                       "Transfer_To_ID_HMI" := "Control_DB".ECnv_Sys[3].Instruction.Transfer_To_ID;
                       "Transfer_From_ID_HMI" := "Control_DB".ECnv_Sys[3].Instruction.Transfer_From_ID;
                       "Pallet_Allignment_HMI" := "Control_DB".ECnv_Sys[3].Instruction.Pallet_Allignment;
                   120603:
                       "Enable_HMI" := "Control_DB".ECnv_Sys[3].Instruction.Enable;
                       "Mode_Change_HMI" := "Control_DB".ECnv_Sys[3].Instruction.Mode_Change;
                       "Task_ID_HMI" := "Control_DB".ECnv_Sys[3].Instruction.Task_ID;
                       "Transfer_To_ID_HMI" := "Control_DB".ECnv_Sys[3].Instruction.Transfer_To_ID;
                       "Transfer_From_ID_HMI" := "Control_DB".ECnv_Sys[3].Instruction.Transfer_From_ID;
                       "Pallet_Allignment_HMI" := "Control_DB".ECnv_Sys[3].Instruction.Pallet_Allignment;
                   120703:
                       "Enable_HMI" := "Control_DB".ECnv_Sys[3].Instruction.Enable;
                       "Mode_Change_HMI" := "Control_DB".ECnv_Sys[3].Instruction.Mode_Change;
                       "Task_ID_HMI" := "Control_DB".ECnv_Sys[3].Instruction.Task_ID;
                       "Transfer_To_ID_HMI" := "Control_DB".ECnv_Sys[3].Instruction.Transfer_To_ID;
                       "Transfer_From_ID_HMI" := "Control_DB".ECnv_Sys[3].Instruction.Transfer_From_ID;
                       "Pallet_Allignment_HMI" := "Control_DB".ECnv_Sys[3].Instruction.Pallet_Allignment;
                   120803:
                       "Enable_HMI" := "Control_DB".ECnv_Sys[3].Instruction.Enable;
                       "Mode_Change_HMI" := "Control_DB".ECnv_Sys[3].Instruction.Mode_Change;
                       "Task_ID_HMI" := "Control_DB".ECnv_Sys[3].Instruction.Task_ID;
                       "Transfer_To_ID_HMI" := "Control_DB".ECnv_Sys[3].Instruction.Transfer_To_ID;
                       "Transfer_From_ID_HMI" := "Control_DB".ECnv_Sys[3].Instruction.Transfer_From_ID;
                       "Pallet_Allignment_HMI" := "Control_DB".ECnv_Sys[3].Instruction.Pallet_Allignment;

                       //SYSTEM 4
                   120004:
                       "Enable_HMI" := "Control_DB".ECnv_Sys[4].Instruction.Enable;
                       "Mode_Change_HMI" := "Control_DB".ECnv_Sys[4].Instruction.Mode_Change;
                       "Task_ID_HMI" := "Control_DB".ECnv_Sys[4].Instruction.Task_ID;
                       "Transfer_To_ID_HMI" := "Control_DB".ECnv_Sys[4].Instruction.Transfer_To_ID;
                       "Transfer_From_ID_HMI" := "Control_DB".ECnv_Sys[4].Instruction.Transfer_From_ID;
                       "Pallet_Allignment_HMI" := "Control_DB".ECnv_Sys[3].Instruction.Pallet_Allignment;
                   120104:
                       "Enable_HMI" := "Control_DB".ECnv_Sys[4].Instruction.Enable;
                       "Mode_Change_HMI" := "Control_DB".ECnv_Sys[4].Instruction.Mode_Change;
                       "Task_ID_HMI" := "Control_DB".ECnv_Sys[4].Instruction.Task_ID;
                       "Transfer_To_ID_HMI" := "Control_DB".ECnv_Sys[4].Instruction.Transfer_To_ID;
                       "Transfer_From_ID_HMI" := "Control_DB".ECnv_Sys[4].Instruction.Transfer_From_ID;
                       "Pallet_Allignment_HMI" := "Control_DB".ECnv_Sys[3].Instruction.Pallet_Allignment;
                   120204:
                       "Enable_HMI" := "Control_DB".ECnv_Sys[4].Instruction.Enable;
                       "Mode_Change_HMI" := "Control_DB".ECnv_Sys[4].Instruction.Mode_Change;
                       "Task_ID_HMI" := "Control_DB".ECnv_Sys[4].Instruction.Task_ID;
                       "Transfer_To_ID_HMI" := "Control_DB".ECnv_Sys[4].Instruction.Transfer_To_ID;
                       "Transfer_From_ID_HMI" := "Control_DB".ECnv_Sys[4].Instruction.Transfer_From_ID;
                       "Pallet_Allignment_HMI" := "Control_DB".ECnv_Sys[3].Instruction.Pallet_Allignment;
                   120304:
                       "Enable_HMI" := "Control_DB".ECnv_Sys[4].Instruction.Enable;
                       "Mode_Change_HMI" := "Control_DB".ECnv_Sys[4].Instruction.Mode_Change;
                       "Task_ID_HMI" := "Control_DB".ECnv_Sys[4].Instruction.Task_ID;
                       "Transfer_To_ID_HMI" := "Control_DB".ECnv_Sys[4].Instruction.Transfer_To_ID;
                       "Transfer_From_ID_HMI" := "Control_DB".ECnv_Sys[4].Instruction.Transfer_From_ID;
                       "Pallet_Allignment_HMI" := "Control_DB".ECnv_Sys[3].Instruction.Pallet_Allignment;
                   120404:
                       "Enable_HMI" := "Control_DB".ECnv_Sys[4].Instruction.Enable;
                       "Mode_Change_HMI" := "Control_DB".ECnv_Sys[4].Instruction.Mode_Change;
                       "Task_ID_HMI" := "Control_DB".ECnv_Sys[4].Instruction.Task_ID;
                       "Transfer_To_ID_HMI" := "Control_DB".ECnv_Sys[4].Instruction.Transfer_To_ID;
                       "Transfer_From_ID_HMI" := "Control_DB".ECnv_Sys[4].Instruction.Transfer_From_ID;
                       "Pallet_Allignment_HMI" := "Control_DB".ECnv_Sys[3].Instruction.Pallet_Allignment;
                   120504:
                       "Enable_HMI" := "Control_DB".ECnv_Sys[4].Instruction.Enable;
                       "Mode_Change_HMI" := "Control_DB".ECnv_Sys[4].Instruction.Mode_Change;
                       "Task_ID_HMI" := "Control_DB".ECnv_Sys[4].Instruction.Task_ID;
                       "Transfer_To_ID_HMI" := "Control_DB".ECnv_Sys[4].Instruction.Transfer_To_ID;
                       "Transfer_From_ID_HMI" := "Control_DB".ECnv_Sys[4].Instruction.Transfer_From_ID;
                       "Pallet_Allignment_HMI" := "Control_DB".ECnv_Sys[3].Instruction.Pallet_Allignment;
                   120604:
                       "Enable_HMI" := "Control_DB".ECnv_Sys[4].Instruction.Enable;
                       "Mode_Change_HMI" := "Control_DB".ECnv_Sys[4].Instruction.Mode_Change;
                       "Task_ID_HMI" := "Control_DB".ECnv_Sys[4].Instruction.Task_ID;
                       "Transfer_To_ID_HMI" := "Control_DB".ECnv_Sys[4].Instruction.Transfer_To_ID;
                       "Transfer_From_ID_HMI" := "Control_DB".ECnv_Sys[4].Instruction.Transfer_From_ID;
                       "Pallet_Allignment_HMI" := "Control_DB".ECnv_Sys[3].Instruction.Pallet_Allignment;
                   120704:
                       "Enable_HMI" := "Control_DB".ECnv_Sys[4].Instruction.Enable;
                       "Mode_Change_HMI" := "Control_DB".ECnv_Sys[4].Instruction.Mode_Change;
                       "Task_ID_HMI" := "Control_DB".ECnv_Sys[4].Instruction.Task_ID;
                       "Transfer_To_ID_HMI" := "Control_DB".ECnv_Sys[4].Instruction.Transfer_To_ID;
                       "Transfer_From_ID_HMI" := "Control_DB".ECnv_Sys[4].Instruction.Transfer_From_ID;
                       "Pallet_Allignment_HMI" := "Control_DB".ECnv_Sys[3].Instruction.Pallet_Allignment;
                   120804:
                       "Enable_HMI" := "Control_DB".ECnv_Sys[4].Instruction.Enable;
                       "Mode_Change_HMI" := "Control_DB".ECnv_Sys[4].Instruction.Mode_Change;
                       "Task_ID_HMI" := "Control_DB".ECnv_Sys[4].Instruction.Task_ID;
                       "Transfer_To_ID_HMI" := "Control_DB".ECnv_Sys[4].Instruction.Transfer_To_ID;
                       "Transfer_From_ID_HMI" := "Control_DB".ECnv_Sys[4].Instruction.Transfer_From_ID;
                       "Pallet_Allignment_HMI" := "Control_DB".ECnv_Sys[3].Instruction.Pallet_Allignment;
                   //SYSTEM 5
                   120005:
                       "Enable_HMI" := "Control_DB".ECnv_Sys[5].Instruction.Enable;
                       "Mode_Change_HMI" := "Control_DB".ECnv_Sys[5].Instruction.Mode_Change;
                       "Task_ID_HMI" := "Control_DB".ECnv_Sys[5].Instruction.Task_ID;
                       "Transfer_To_ID_HMI" := "Control_DB".ECnv_Sys[5].Instruction.Transfer_To_ID;
                       "Transfer_From_ID_HMI" := "Control_DB".ECnv_Sys[5].Instruction.Transfer_From_ID;
                       "Pallet_Allignment_HMI" := "Control_DB".ECnv_Sys[5].Instruction.Pallet_Allignment;
                   120105:
                       "Enable_HMI" := "Control_DB".ECnv_Sys[5].Instruction.Enable;
                       "Mode_Change_HMI" := "Control_DB".ECnv_Sys[5].Instruction.Mode_Change;
                       "Task_ID_HMI" := "Control_DB".ECnv_Sys[5].Instruction.Task_ID;
                       "Transfer_To_ID_HMI" := "Control_DB".ECnv_Sys[5].Instruction.Transfer_To_ID;
                       "Transfer_From_ID_HMI" := "Control_DB".ECnv_Sys[5].Instruction.Transfer_From_ID;
                       "Pallet_Allignment_HMI" := "Control_DB".ECnv_Sys[5].Instruction.Pallet_Allignment;
                   120205:
                       "Enable_HMI" := "Control_DB".ECnv_Sys[5].Instruction.Enable;
                       "Mode_Change_HMI" := "Control_DB".ECnv_Sys[5].Instruction.Mode_Change;
                       "Task_ID_HMI" := "Control_DB".ECnv_Sys[5].Instruction.Task_ID;
                       "Transfer_To_ID_HMI" := "Control_DB".ECnv_Sys[5].Instruction.Transfer_To_ID;
                       "Transfer_From_ID_HMI" := "Control_DB".ECnv_Sys[5].Instruction.Transfer_From_ID;
                       "Pallet_Allignment_HMI" := "Control_DB".ECnv_Sys[5].Instruction.Pallet_Allignment;
                   120305:
                       "Enable_HMI" := "Control_DB".ECnv_Sys[5].Instruction.Enable;
                       "Mode_Change_HMI" := "Control_DB".ECnv_Sys[5].Instruction.Mode_Change;
                       "Task_ID_HMI" := "Control_DB".ECnv_Sys[5].Instruction.Task_ID;
                       "Transfer_To_ID_HMI" := "Control_DB".ECnv_Sys[5].Instruction.Transfer_To_ID;
                       "Transfer_From_ID_HMI" := "Control_DB".ECnv_Sys[5].Instruction.Transfer_From_ID;
                       "Pallet_Allignment_HMI" := "Control_DB".ECnv_Sys[5].Instruction.Pallet_Allignment;
                   120405:
                       "Enable_HMI" := "Control_DB".ECnv_Sys[5].Instruction.Enable;
                       "Mode_Change_HMI" := "Control_DB".ECnv_Sys[5].Instruction.Mode_Change;
                       "Task_ID_HMI" := "Control_DB".ECnv_Sys[5].Instruction.Task_ID;
                       "Transfer_To_ID_HMI" := "Control_DB".ECnv_Sys[5].Instruction.Transfer_To_ID;
                       "Transfer_From_ID_HMI" := "Control_DB".ECnv_Sys[5].Instruction.Transfer_From_ID;
                       "Pallet_Allignment_HMI" := "Control_DB".ECnv_Sys[5].Instruction.Pallet_Allignment;
                   120505:
                       "Enable_HMI" := "Control_DB".ECnv_Sys[5].Instruction.Enable;
                       "Mode_Change_HMI" := "Control_DB".ECnv_Sys[5].Instruction.Mode_Change;
                       "Task_ID_HMI" := "Control_DB".ECnv_Sys[5].Instruction.Task_ID;
                       "Transfer_To_ID_HMI" := "Control_DB".ECnv_Sys[5].Instruction.Transfer_To_ID;
                       "Transfer_From_ID_HMI" := "Control_DB".ECnv_Sys[5].Instruction.Transfer_From_ID;
                       "Pallet_Allignment_HMI" := "Control_DB".ECnv_Sys[5].Instruction.Pallet_Allignment;
                   120605:
                       "Enable_HMI" := "Control_DB".ECnv_Sys[5].Instruction.Enable;
                       "Mode_Change_HMI" := "Control_DB".ECnv_Sys[5].Instruction.Mode_Change;
                       "Task_ID_HMI" := "Control_DB".ECnv_Sys[5].Instruction.Task_ID;
                       "Transfer_To_ID_HMI" := "Control_DB".ECnv_Sys[5].Instruction.Transfer_To_ID;
                       "Transfer_From_ID_HMI" := "Control_DB".ECnv_Sys[5].Instruction.Transfer_From_ID;
                       "Pallet_Allignment_HMI" := "Control_DB".ECnv_Sys[5].Instruction.Pallet_Allignment;
                   120705:
                       "Enable_HMI" := "Control_DB".ECnv_Sys[5].Instruction.Enable;
                       "Mode_Change_HMI" := "Control_DB".ECnv_Sys[5].Instruction.Mode_Change;
                       "Task_ID_HMI" := "Control_DB".ECnv_Sys[5].Instruction.Task_ID;
                       "Transfer_To_ID_HMI" := "Control_DB".ECnv_Sys[5].Instruction.Transfer_To_ID;
                       "Transfer_From_ID_HMI" := "Control_DB".ECnv_Sys[5].Instruction.Transfer_From_ID;
                       "Pallet_Allignment_HMI" := "Control_DB".ECnv_Sys[5].Instruction.Pallet_Allignment;
                   120805:
                       "Enable_HMI" := "Control_DB".ECnv_Sys[5].Instruction.Enable;
                       "Mode_Change_HMI" := "Control_DB".ECnv_Sys[5].Instruction.Mode_Change;
                       "Task_ID_HMI" := "Control_DB".ECnv_Sys[5].Instruction.Task_ID;
                       "Transfer_To_ID_HMI" := "Control_DB".ECnv_Sys[5].Instruction.Transfer_To_ID;
                       "Transfer_From_ID_HMI" := "Control_DB".ECnv_Sys[5].Instruction.Transfer_From_ID;
                       "Pallet_Allignment_HMI" := "Control_DB".ECnv_Sys[5].Instruction.Pallet_Allignment;
               END_CASE;
               // "Screen_DB".Charge_Cnv_Commands := 0;
           END_IF;
       END_REGION

       REGION CHARGE DATA FROM HMI (AFTER CHARGE DATA)
           IF NOT "Screen_DB".Charge_Cnv_Commands AND "HMI_DB".ScreenNo_Main = 2 AND NOT #R_Charge_Cnv_Commands.Q THEN
               CASE "CNV_ID_HMI" OF
                       //SYSTEM 1
                   120101:
                       "Feed_ECNV"(System_No := 1,
                                   Safety_OK:="Remote_Panel_DB_1".Safety_OK,
                                   Overhang_Left:="CVTD1 OVERHANG LEFT",
                                   Overhang_Right:="CVTD1 OVERHANG RIGHT",
                                   System_Busy:="System_1_Busy");
                   120201:
                       "Feed_ECNV"(System_No := 1,
                                   Safety_OK:="Remote_Panel_DB_1".Safety_OK,
                                   Overhang_Left:="CVTD1 OVERHANG LEFT",
                                   Overhang_Right:="CVTD1 OVERHANG RIGHT",
                                   System_Busy:="System_1_Busy");
                   120301:
                       "Feed_ECNV"(System_No := 1,
                                   Safety_OK:="Remote_Panel_DB_1".Safety_OK,
                                   Overhang_Left:="CVTD1 OVERHANG LEFT",
                                   Overhang_Right:="CVTD1 OVERHANG RIGHT",
                                   System_Busy:="System_1_Busy");
                   120401:
                       "Feed_ECNV"(System_No := 1,
                                   Safety_OK:="Remote_Panel_DB_1".Safety_OK,
                                   Overhang_Left:="CVTD1 OVERHANG LEFT",
                                   Overhang_Right:="CVTD1 OVERHANG RIGHT",
                                   System_Busy:="System_1_Busy");
                   120501:
                       "Feed_ECNV"(System_No := 1,
                                   Safety_OK:="Remote_Panel_DB_1".Safety_OK,
                                   Overhang_Left:="CVTD1 OVERHANG LEFT",
                                   Overhang_Right:="CVTD1 OVERHANG RIGHT",
                                   System_Busy:="System_1_Busy");
                   120601:
                       "Feed_ECNV"(System_No := 1,
                                   Safety_OK:="Remote_Panel_DB_1".Safety_OK,
                                   Overhang_Left:="CVTD1 OVERHANG LEFT",
                                   Overhang_Right:="CVTD1 OVERHANG RIGHT",
                                   System_Busy:="System_1_Busy");
                   120701:
                       "Feed_ECNV"(System_No := 1,
                                   Safety_OK:="Remote_Panel_DB_1".Safety_OK,
                                   Overhang_Left:="CVTD1 OVERHANG LEFT",
                                   Overhang_Right:="CVTD1 OVERHANG RIGHT",
                                   System_Busy:="System_1_Busy");
                   120801:
                       "Feed_ECNV"(System_No := 1,
                                   Safety_OK:="Remote_Panel_DB_1".Safety_OK,
                                   Overhang_Left:="CVTD1 OVERHANG LEFT",
                                   Overhang_Right:="CVTD1 OVERHANG RIGHT",
                                   System_Busy:="System_1_Busy");

                       //SYSTEM 2
                   120102:
                       "Feed_ECNV"(System_No := 2,
                                   Safety_OK:="Remote_Panel_DB_2".Safety_OK,
                                   Overhang_Left:="CVTD2 OVERHANG LEFT",
                                   Overhang_Right:="CVTD2 OVERHANG RIGHT",
                                   System_Busy:="System_2_Busy");
                   120202:
                       "Feed_ECNV"(System_No := 2,
                                   Safety_OK:="Remote_Panel_DB_2".Safety_OK,
                                   Overhang_Left:="CVTD2 OVERHANG LEFT",
                                   Overhang_Right:="CVTD2 OVERHANG RIGHT",
                                   System_Busy:="System_2_Busy");
                   120302:
                       "Feed_ECNV"(System_No := 2,
                                   Safety_OK:="Remote_Panel_DB_2".Safety_OK,
                                   Overhang_Left:="CVTD2 OVERHANG LEFT",
                                   Overhang_Right:="CVTD2 OVERHANG RIGHT",
                                   System_Busy:="System_2_Busy");
                   120402:
                       "Feed_ECNV"(System_No := 2,
                                   Safety_OK:="Remote_Panel_DB_2".Safety_OK,
                                   Overhang_Left:="CVTD2 OVERHANG LEFT",
                                   Overhang_Right:="CVTD2 OVERHANG RIGHT",
                                   System_Busy:="System_2_Busy");
                   120502:
                       "Feed_ECNV"(System_No := 2,
                                   Safety_OK:="Remote_Panel_DB_2".Safety_OK,
                                   Overhang_Left:="CVTD2 OVERHANG LEFT",
                                   Overhang_Right:="CVTD2 OVERHANG RIGHT",
                                   System_Busy:="System_2_Busy");
                   120602:
                       "Feed_ECNV"(System_No := 2,
                                   Safety_OK:="Remote_Panel_DB_2".Safety_OK,
                                   Overhang_Left:="CVTD2 OVERHANG LEFT",
                                   Overhang_Right:="CVTD2 OVERHANG RIGHT",
                                   System_Busy:="System_2_Busy");
                   120702:
                       "Feed_ECNV"(System_No := 2,
                                   Safety_OK:="Remote_Panel_DB_2".Safety_OK,
                                   Overhang_Left:="CVTD2 OVERHANG LEFT",
                                   Overhang_Right:="CVTD2 OVERHANG RIGHT",
                                   System_Busy:="System_2_Busy");
                   120802:
                       "Feed_ECNV"(System_No := 2,
                                   Safety_OK:="Remote_Panel_DB_2".Safety_OK,
                                   Overhang_Left:="CVTD2 OVERHANG LEFT",
                                   Overhang_Right:="CVTD2 OVERHANG RIGHT",
                                   System_Busy:="System_2_Busy");

                       //SYSTEM 3
                   120103:
                       "Feed_ECNV"(System_No := 3,
                                   Safety_OK:="Remote_Panel_DB_3".Safety_OK,
                                   Overhang_Left:="CVTD3 OVERHANG LEFT",
                                   Overhang_Right:="CVTD3 OVERHANG RIGHT",
                                   System_Busy:="System_3_Busy");
                   120203:
                       "Feed_ECNV"(System_No := 3,
                                   Safety_OK:="Remote_Panel_DB_3".Safety_OK,
                                   Overhang_Left:="CVTD3 OVERHANG LEFT",
                                   Overhang_Right:="CVTD3 OVERHANG RIGHT",
                                   System_Busy:="System_3_Busy");
                   120303:
                       "Feed_ECNV"(System_No := 3,
                                   Safety_OK:="Remote_Panel_DB_3".Safety_OK,
                                   Overhang_Left:="CVTD3 OVERHANG LEFT",
                                   Overhang_Right:="CVTD3 OVERHANG RIGHT",
                                   System_Busy:="System_3_Busy");
                   120403:
                       "Feed_ECNV"(System_No := 3,
                                   Safety_OK:="Remote_Panel_DB_3".Safety_OK,
                                   Overhang_Left:="CVTD3 OVERHANG LEFT",
                                   Overhang_Right:="CVTD3 OVERHANG RIGHT",
                                   System_Busy:="System_3_Busy");
                   120503:
                       "Feed_ECNV"(System_No := 3,
                                   Safety_OK:="Remote_Panel_DB_3".Safety_OK,
                                   Overhang_Left:="CVTD3 OVERHANG LEFT",
                                   Overhang_Right:="CVTD3 OVERHANG RIGHT",
                                   System_Busy:="System_3_Busy");
                   120603:
                       "Feed_ECNV"(System_No := 3,
                                   Safety_OK:="Remote_Panel_DB_3".Safety_OK,
                                   Overhang_Left:="CVTD3 OVERHANG LEFT",
                                   Overhang_Right:="CVTD3 OVERHANG RIGHT",
                                   System_Busy:="System_3_Busy");
                   120703:
                       "Feed_ECNV"(System_No := 3,
                                   Safety_OK:="Remote_Panel_DB_3".Safety_OK,
                                   Overhang_Left:="CVTD3 OVERHANG LEFT",
                                   Overhang_Right:="CVTD3 OVERHANG RIGHT",
                                   System_Busy:="System_3_Busy");
                   120803:
                       "Feed_ECNV"(System_No := 3,
                                   Safety_OK:="Remote_Panel_DB_3".Safety_OK,
                                   Overhang_Left:="CVTD3 OVERHANG LEFT",
                                   Overhang_Right:="CVTD3 OVERHANG RIGHT",
                                   System_Busy:="System_3_Busy");

                       //SYSTEM 4
                   120104:
                       "Feed_ECNV"(System_No := 4,
                                   Safety_OK:="Remote_Panel_DB_4".Safety_OK,
                                   Overhang_Left:="CVTD4 OVERHANG LEFT",
                                   Overhang_Right:="CVTD4 OVERHANG RIGHT",
                                   System_Busy:="System_4_Busy");
                   120204:
                       "Feed_ECNV"(System_No := 4,
                                   Safety_OK:="Remote_Panel_DB_4".Safety_OK,
                                   Overhang_Left:="CVTD4 OVERHANG LEFT",
                                   Overhang_Right:="CVTD4 OVERHANG RIGHT",
                                   System_Busy:="System_4_Busy");
                   120304:
                       "Feed_ECNV"(System_No := 4,
                                   Safety_OK:="Remote_Panel_DB_4".Safety_OK,
                                   Overhang_Left:="CVTD4 OVERHANG LEFT",
                                   Overhang_Right:="CVTD4 OVERHANG RIGHT",
                                   System_Busy:="System_4_Busy");
                   120404:
                       "Feed_ECNV"(System_No := 4,
                                   Safety_OK:="Remote_Panel_DB_4".Safety_OK,
                                   Overhang_Left:="CVTD4 OVERHANG LEFT",
                                   Overhang_Right:="CVTD4 OVERHANG RIGHT",
                                   System_Busy:="System_4_Busy");
                   120504:
                       "Feed_ECNV"(System_No := 4,
                                   Safety_OK:="Remote_Panel_DB_4".Safety_OK,
                                   Overhang_Left:="CVTD4 OVERHANG LEFT",
                                   Overhang_Right:="CVTD4 OVERHANG RIGHT",
                                   System_Busy:="System_4_Busy");
                   120604:
                       "Feed_ECNV"(System_No := 4,
                                   Safety_OK:="Remote_Panel_DB_4".Safety_OK,
                                   Overhang_Left:="CVTD4 OVERHANG LEFT",
                                   Overhang_Right:="CVTD4 OVERHANG RIGHT",
                                   System_Busy:="System_4_Busy");
                   120704:
                       "Feed_ECNV"(System_No := 4,
                                   Safety_OK:="Remote_Panel_DB_4".Safety_OK,
                                   Overhang_Left:="CVTD4 OVERHANG LEFT",
                                   Overhang_Right:="CVTD4 OVERHANG RIGHT",
                                   System_Busy:="System_4_Busy");
                   120804:
                       "Feed_ECNV"(System_No := 4,
                                   Safety_OK:="Remote_Panel_DB_4".Safety_OK,
                                   Overhang_Left:="CVTD4 OVERHANG LEFT",
                                   Overhang_Right:="CVTD4 OVERHANG RIGHT",
                                   System_Busy:="System_4_Busy");

                       //SYSTEM 5
                   120105:
                       "Feed_ECNV"(System_No := 5,
                                   Safety_OK:="Remote_Panel_DB_5".Safety_OK,
                                   Overhang_Left:="CVTD5 OVERHANG LEFT",
                                   Overhang_Right:="CVTD5 OVERHANG RIGHT",
                                   System_Busy:="System_5_Busy");
                   120205:
                       "Feed_ECNV"(System_No := 5,
                                   Safety_OK:="Remote_Panel_DB_5".Safety_OK,
                                   Overhang_Left:="CVTD5 OVERHANG LEFT",
                                   Overhang_Right:="CVTD5 OVERHANG RIGHT",
                                   System_Busy:="System_5_Busy");
                   120305:
                       "Feed_ECNV"(System_No := 5,
                                   Safety_OK:="Remote_Panel_DB_5".Safety_OK,
                                   Overhang_Left:="CVTD5 OVERHANG LEFT",
                                   Overhang_Right:="CVTD5 OVERHANG RIGHT",
                                   System_Busy:="System_5_Busy");
                   120405:
                       "Feed_ECNV"(System_No := 5,
                                   Safety_OK:="Remote_Panel_DB_5".Safety_OK,
                                   Overhang_Left:="CVTD5 OVERHANG LEFT",
                                   Overhang_Right:="CVTD5 OVERHANG RIGHT",
                                   System_Busy:="System_5_Busy");
                   120505:
                       "Feed_ECNV"(System_No := 5,
                                   Safety_OK:="Remote_Panel_DB_5".Safety_OK,
                                   Overhang_Left:="CVTD5 OVERHANG LEFT",
                                   Overhang_Right:="CVTD5 OVERHANG RIGHT",
                                   System_Busy:="System_5_Busy");
                   120605:
                       "Feed_ECNV"(System_No := 5,
                                   Safety_OK:="Remote_Panel_DB_5".Safety_OK,
                                   Overhang_Left:="CVTD5 OVERHANG LEFT",
                                   Overhang_Right:="CVTD5 OVERHANG RIGHT",
                                   System_Busy:="System_5_Busy");
                   120705:
                       "Feed_ECNV"(System_No := 5,
                                   Safety_OK:="Remote_Panel_DB_5".Safety_OK,
                                   Overhang_Left:="CVTD5 OVERHANG LEFT",
                                   Overhang_Right:="CVTD5 OVERHANG RIGHT",
                                   System_Busy:="System_5_Busy");
                   120805:
                       "Feed_ECNV"(System_No := 5,
                                   Safety_OK:="Remote_Panel_DB_5".Safety_OK,
                                   Overhang_Left:="CVTD5 OVERHANG LEFT",
                                   Overhang_Right:="CVTD5 OVERHANG RIGHT",
                                   System_Busy:="System_5_Busy");
               END_CASE;
           END_IF;
       END_REGION
   END_REGION

   REGION Assign Conveyor 2
       REGION CHARGE DATA FROM THE CORRECT CONVEYOR
           //CHARGE DATA CHANGING CONVEYORS ID
           IF "CNV_ID_HMI(1)" <> "CNV_ID_HM_Old(1)" THEN
               "Screen_DB".Charge_Cnv_Commands := TRUE;
               "CNV_ID_HM_Old(1)" := "CNV_ID_HMI(1)";
           END_IF;
           #R_Charge_Cnv_Commands(CLK := "Screen_DB".Charge_Cnv_Commands OR "HMI_DB".ScreenNo_Main = 2);

